TYPE ET_ContourType_1 :
(
	ET_ContourType_eNone := 0,
	ET_ContourType_eCircle := 1,
	ET_ContourType_eEllipse := 2,
	ET_ContourType_eSquare := 3
);
END_TYPE

(* stored: Version 1.1.0.1, ProductVersion 3.1.4024.15
   DUT ET_ContourType_1: Id {6732b04c-19a0-4c4a-a710-44e20da8f46a} *)
